(* IEC 61131-3 sources: plc-process-lib/tests/POUs/Suites/FB_Valve_Test (part 2) *)

(* ---- PowerLossStopsWithoutFault.method.impl.st ---- *)
coUnit.TEST('Valve_PowerLoss_StopsWithoutFault');

stCfg.tTravel := T#10S;
fbVlv.xZsc := TRUE;
fbVlv(itfTime := fbTime, stCmd := stCmd, stRetain := stRetain, stCfg := stCfg);
stCmd.xOpen := TRUE;
fbVlv(itfTime := fbTime, stCmd := stCmd, stRetain := stRetain, stCfg := stCfg);
fbVlv.xZsc := FALSE;
FOR iStep := 1 TO 10 DO
    fbTime.Advance(tStep := T#100MS);
    fbVlv(itfTime := fbTime, stCmd := stCmd, stRetain := stRetain, stCfg := stCfg);
END_FOR
fbVlv.xPowerOk := FALSE;
fbTime.Advance(tStep := T#100MS);
fbVlv(itfTime := fbTime, stCmd := stCmd, stRetain := stRetain, stCfg := stCfg);
AssertTrue(Condition := fbVlv.stSts.eState = E_ValveState.Intermediate, Message := 'Intermediate on power loss');
AssertFalse(Condition := fbVlv.xQOpen, Message := 'output off');
AssertEquals_WORD(Expected := GVL_Const.VLV_WRN_POWER_LOST,
                  Actual := fbVlv.stSts.stCommon.wWarning AND GVL_Const.VLV_WRN_POWER_LOST, Message := 'POWER_LOST');
AssertEquals_WORD(Expected := 0, Actual := fbVlv.stSts.stCommon.wFault, Message := 'no fault');
AssertFalse(Condition := fbVlv.Fault, Message := 'not Fault');
stCmd.xOpen := TRUE;
fbTime.Advance(tStep := T#100MS);
fbVlv(itfTime := fbTime, stCmd := stCmd, stRetain := stRetain, stCfg := stCfg);
AssertTrue(Condition := fbVlv.stSts.stCommon.eCmdResult = E_CmdResult.RejectedInhibit,
           Message := 'command without power: RejectedInhibit');
FOR iStep := 1 TO 120 DO                                                // 12 с без напряжения
    fbTime.Advance(tStep := T#100MS);
    fbVlv(itfTime := fbTime, stCmd := stCmd, stRetain := stRetain, stCfg := stCfg);
END_FOR
AssertEquals_WORD(Expected := 0, Actual := fbVlv.stSts.stCommon.wFault, Message := 'travel supervision suspended');
fbVlv.xPowerOk := TRUE;
fbTime.Advance(tStep := T#100MS);
fbVlv(itfTime := fbTime, stCmd := stCmd, stRetain := stRetain, stCfg := stCfg);
AssertTrue(Condition := fbVlv.stSts.eState = E_ValveState.Intermediate, Message := 'Manual stays: target cleared');
AssertFalse(Condition := fbVlv.xQOpen, Message := 'no output in Manual');
stCmd.stCommon.xSetAuto := TRUE;
fbVlv.xAutoOpen := TRUE;
fbTime.Advance(tStep := T#100MS);
fbVlv(itfTime := fbTime, stCmd := stCmd, stRetain := stRetain, stCfg := stCfg);
AssertTrue(Condition := fbVlv.xQOpen, Message := 'Auto drives to target');
AssertTrue(Condition := fbVlv.Available, Message := 'available in Auto with power');
fbVlv.xPowerOk := FALSE;
fbTime.Advance(tStep := T#100MS);
fbVlv(itfTime := fbTime, stCmd := stCmd, stRetain := stRetain, stCfg := stCfg);
AssertFalse(Condition := fbVlv.xQOpen, Message := 'off again without power');
AssertFalse(Condition := fbVlv.Available, Message := 'not available without power');
AssertEquals_WORD(Expected := 0, Actual := fbVlv.stSts.stCommon.wStatus AND GVL_Const.VLV_STS_AVAILABLE,
                  Message := 'AVAILABLE bit off without power');
fbVlv.xPowerOk := TRUE;
fbTime.Advance(tStep := T#100MS);
fbVlv(itfTime := fbTime, stCmd := stCmd, stRetain := stRetain, stCfg := stCfg);
AssertTrue(Condition := fbVlv.xQOpen, Message := 'Auto resumes after power returns');
AssertTrue(Condition := fbVlv.stSts.eState = E_ValveState.Opening, Message := 'Opening');

coUnit.TEST_FINISHED();

(* ---- ResetCauseClearsWithinWindowFaultCleared.method.decl.st ---- *)
// TorqueTrip, Reset при сработавшей муфте: отказ держится; муфта отпустила через 1 с — отказ снят в окне
// tResetWindow без второго результата (и после конца окна RejectedFault нет).
METHOD PRIVATE ResetCauseClearsWithinWindowFaultCleared
VAR
    fbTime   : FB_FakeTime;       // подменное время, старт 1 ч
    fbVlv    : FB_Valve;          // арматура под тестом
    stCmd    : ST_ValveCmd;       // команды HMI
    stRetain : ST_DeviceRetain;   // режим Manual по умолчанию, счётчики
    stCfg    : ST_ValveCfg;       // конфигурация (умолчания: Motorized, ZSO и ZSC)
    iStep    : INT;               // шаг цикла
    uiSeq    : UINT;              // номер команды после Reset
END_VAR

(* ---- ResetCauseClearsWithinWindowFaultCleared.method.impl.st ---- *)
coUnit.TEST('Valve_Reset_CauseClearsWithinWindow_FaultCleared');

stCfg.xTorqueUsed := TRUE;
fbVlv.xZsc := TRUE;
fbVlv(itfTime := fbTime, stCmd := stCmd, stRetain := stRetain, stCfg := stCfg);
stCmd.xOpen := TRUE;
fbVlv(itfTime := fbTime, stCmd := stCmd, stRetain := stRetain, stCfg := stCfg);
fbVlv.xZsc := FALSE;
FOR iStep := 1 TO 10 DO
    fbTime.Advance(tStep := T#100MS);
    fbVlv(itfTime := fbTime, stCmd := stCmd, stRetain := stRetain, stCfg := stCfg);
END_FOR
fbVlv.xTorqueOpen := TRUE;
fbTime.Advance(tStep := T#100MS);
fbVlv(itfTime := fbTime, stCmd := stCmd, stRetain := stRetain, stCfg := stCfg);
AssertEquals_WORD(Expected := GVL_Const.VLV_FLT_TORQUE_TRIP, Actual := fbVlv.stSts.stCommon.wFault,
                  Message := 'TorqueTrip');
stCmd.stCommon.xReset := TRUE;
// t1: Reset, муфта сработана
fbVlv(itfTime := fbTime, stCmd := stCmd, stRetain := stRetain, stCfg := stCfg);
uiSeq := fbVlv.stSts.stCommon.uiCmdSeq;
AssertEquals_WORD(Expected := GVL_Const.VLV_FLT_TORQUE_TRIP, Actual := fbVlv.stSts.stCommon.wFault,
                  Message := 'cause active right after Reset');
FOR iStep := 1 TO 9 DO                                                  // t1 + 0,9 с
    fbTime.Advance(tStep := T#100MS);
    fbVlv(itfTime := fbTime, stCmd := stCmd, stRetain := stRetain, stCfg := stCfg);
END_FOR
AssertEquals_WORD(Expected := GVL_Const.VLV_FLT_TORQUE_TRIP, Actual := fbVlv.stSts.stCommon.wFault,
                  Message := 'still faulted while torque is on');
fbVlv.xTorqueOpen := FALSE;
fbTime.Advance(tStep := T#100MS);
// t1 + 1,0 с: муфта отпустила
fbVlv(itfTime := fbTime, stCmd := stCmd, stRetain := stRetain, stCfg := stCfg);
AssertEquals_WORD(Expected := 0, Actual := fbVlv.stSts.stCommon.wFault, Message := 'cleared within the window');
FOR iStep := 1 TO 30 DO                                                 // дальше конца окна
    fbTime.Advance(tStep := T#100MS);
    fbVlv(itfTime := fbTime, stCmd := stCmd, stRetain := stRetain, stCfg := stCfg);
END_FOR
AssertEquals_UINT(Expected := uiSeq, Actual := fbVlv.stSts.stCommon.uiCmdSeq, Message := 'no second result');
AssertTrue(Condition := fbVlv.stSts.stCommon.eCmdResult = E_CmdResult.Accepted, Message := 'last result Accepted');
AssertFalse(Condition := fbVlv.xQOpen, Message := 'no restart in Manual');

coUnit.TEST_FINISHED();

(* ---- ReverseAfterEndStopWaitsReversePause.method.decl.st ---- *)
// Motorized: ход на открытие дошёл до ZSO на t1 (выход «открывать» снят), сразу команда «закрыть»:
// выход «закрывать» не включается, пока от снятия «открывать» не прошла пауза tReverse = 1 с (на
// t1 + 0,9 с — ещё нет), ровно на t1 + 1,0 с — Closing. То же после стопа в ходе на закрытие (t2) и
// команды «открыть» через 0,2 с: «открывать» включается только на t2 + 1,0 с. Двигатель на выбеге
// встречным включением не реверсируется, даже если ход перед этим остановил концевик или стоп.
METHOD PRIVATE ReverseAfterEndStopWaitsReversePause
VAR
    fbTime   : FB_FakeTime;       // подменное время, старт 1 ч
    fbVlv    : FB_Valve;          // арматура под тестом
    stCmd    : ST_ValveCmd;       // команды HMI
    stRetain : ST_DeviceRetain;   // режим Manual по умолчанию, счётчики
    stCfg    : ST_ValveCfg;       // конфигурация (умолчания: Motorized, ZSO и ZSC, tReverse = 1 с)
    iStep    : INT;               // шаг цикла
    xEverOn  : BOOL;              // выход включался во время паузы
END_VAR

(* ---- ReverseAfterEndStopWaitsReversePause.method.impl.st ---- *)
coUnit.TEST('Valve_ReverseAfterEndStop_WaitsReversePause');

fbVlv.xZsc := TRUE;
// закрыта
fbVlv(itfTime := fbTime, stCmd := stCmd, stRetain := stRetain, stCfg := stCfg);
stCmd.xOpen := TRUE;
fbVlv(itfTime := fbTime, stCmd := stCmd, stRetain := stRetain, stCfg := stCfg);
fbVlv.xZsc := FALSE;
FOR iStep := 1 TO 20 DO                                                 // открывается 2 с
    fbTime.Advance(tStep := T#100MS);
    fbVlv(itfTime := fbTime, stCmd := stCmd, stRetain := stRetain, stCfg := stCfg);
END_FOR
fbVlv.xZso := TRUE;
fbTime.Advance(tStep := T#100MS);
// t1: ZSO, выход «открывать» снят
fbVlv(itfTime := fbTime, stCmd := stCmd, stRetain := stRetain, stCfg := stCfg);
AssertTrue(Condition := fbVlv.stSts.eState = E_ValveState.Open, Message := 'Open on ZSO');
AssertFalse(Condition := fbVlv.xQOpen, Message := 'open contactor off at ZSO');
stCmd.xClose := TRUE;
fbTime.Advance(tStep := T#100MS);
// t1 + 0,1 с: команда «закрыть»
fbVlv(itfTime := fbTime, stCmd := stCmd, stRetain := stRetain, stCfg := stCfg);
AssertTrue(Condition := fbVlv.stSts.stCommon.eCmdResult = E_CmdResult.Accepted, Message := 'close accepted');
xEverOn := fbVlv.xQOpen OR fbVlv.xQClose;
FOR iStep := 1 TO 8 DO                                                  // до t1 + 0,9 с
    fbTime.Advance(tStep := T#100MS);
    fbVlv(itfTime := fbTime, stCmd := stCmd, stRetain := stRetain, stCfg := stCfg);
    xEverOn := xEverOn OR fbVlv.xQOpen OR fbVlv.xQClose;
END_FOR
AssertFalse(Condition := xEverOn, Message := 'no reverse start within tReverse after end stop');
AssertTrue(Condition := fbVlv.stSts.eState = E_ValveState.Open, Message := 'waits at Open');
fbTime.Advance(tStep := T#100MS);
// t1 + 1,0 с
fbVlv(itfTime := fbTime, stCmd := stCmd, stRetain := stRetain, stCfg := stCfg);
AssertTrue(Condition := fbVlv.stSts.eState = E_ValveState.Closing, Message := 'Closing at t1 + tReverse');
AssertTrue(Condition := fbVlv.xQClose, Message := 'close contactor on at t1 + tReverse');
fbVlv.xZso := FALSE;
FOR iStep := 1 TO 20 DO                                                 // закрывается 2 с
    fbTime.Advance(tStep := T#100MS);
    fbVlv(itfTime := fbTime, stCmd := stCmd, stRetain := stRetain, stCfg := stCfg);
END_FOR
stCmd.xStop := TRUE;
// t2: стоп в ходе
fbVlv(itfTime := fbTime, stCmd := stCmd, stRetain := stRetain, stCfg := stCfg);
AssertTrue(Condition := fbVlv.stSts.eState = E_ValveState.Intermediate, Message := 'Intermediate after stop');
stCmd.xOpen := TRUE;
fbTime.Advance(tStep := T#200MS);
// t2 + 0,2 с: команда «открыть»
fbVlv(itfTime := fbTime, stCmd := stCmd, stRetain := stRetain, stCfg := stCfg);
AssertTrue(Condition := fbVlv.stSts.stCommon.eCmdResult = E_CmdResult.Accepted, Message := 'open accepted');
xEverOn := fbVlv.xQOpen OR fbVlv.xQClose;
FOR iStep := 1 TO 7 DO                                                  // до t2 + 0,9 с
    fbTime.Advance(tStep := T#100MS);
    fbVlv(itfTime := fbTime, stCmd := stCmd, stRetain := stRetain, stCfg := stCfg);
    xEverOn := xEverOn OR fbVlv.xQOpen OR fbVlv.xQClose;
END_FOR
AssertFalse(Condition := xEverOn, Message := 'no reverse start within tReverse after stop');
fbTime.Advance(tStep := T#100MS);
// t2 + 1,0 с
fbVlv(itfTime := fbTime, stCmd := stCmd, stRetain := stRetain, stCfg := stCfg);
AssertTrue(Condition := fbVlv.stSts.eState = E_ValveState.Opening, Message := 'Opening at t2 + tReverse');
AssertTrue(Condition := fbVlv.xQOpen, Message := 'open contactor on at t2 + tReverse');

coUnit.TEST_FINISHED();

(* ---- ReversePausesBeforeOppositeDirection.method.decl.st ---- *)
// Motorized открывается; команда «закрыть» в ходе: Reversing, оба выхода сняты на tReverse = 1 с (на
// t1 + 0,9 с ещё сняты), ровно на t1 + 1,0 с включается xQClose.
METHOD PRIVATE ReversePausesBeforeOppositeDirection
VAR
    fbTime   : FB_FakeTime;       // подменное время, старт 1 ч
    fbVlv    : FB_Valve;          // арматура под тестом
    stCmd    : ST_ValveCmd;       // команды HMI
    stRetain : ST_DeviceRetain;   // режим Manual по умолчанию, счётчики
    stCfg    : ST_ValveCfg;       // конфигурация (умолчания: Motorized, ZSO и ZSC)
    iStep    : INT;               // шаг цикла
    xEverOn  : BOOL;              // выход включался во время паузы
END_VAR

(* ---- ReversePausesBeforeOppositeDirection.method.impl.st ---- *)
coUnit.TEST('Valve_Reverse_PausesBeforeOppositeDirection');

fbVlv.xZsc := TRUE;
// закрыта
fbVlv(itfTime := fbTime, stCmd := stCmd, stRetain := stRetain, stCfg := stCfg);
stCmd.xOpen := TRUE;
// Opening
fbVlv(itfTime := fbTime, stCmd := stCmd, stRetain := stRetain, stCfg := stCfg);
fbVlv.xZsc := FALSE;
FOR iStep := 1 TO 20 DO                                                 // открывается 2 с
    fbTime.Advance(tStep := T#100MS);
    fbVlv(itfTime := fbTime, stCmd := stCmd, stRetain := stRetain, stCfg := stCfg);
END_FOR
AssertTrue(Condition := fbVlv.xQOpen, Message := 'opening');
stCmd.xClose := TRUE;
// t1: смена направления
fbVlv(itfTime := fbTime, stCmd := stCmd, stRetain := stRetain, stCfg := stCfg);
AssertTrue(Condition := fbVlv.stSts.eState = E_ValveState.Reversing, Message := 'Reversing on direction change');
AssertFalse(Condition := fbVlv.xQOpen OR fbVlv.xQClose, Message := 'both outputs off during the pause');
AssertTrue(Condition := fbVlv.stSts.stCommon.eCmdResult = E_CmdResult.Accepted, Message := 'close accepted');
FOR iStep := 1 TO 9 DO                                                  // t1 + 0,9 с
    fbTime.Advance(tStep := T#100MS);
    fbVlv(itfTime := fbTime, stCmd := stCmd, stRetain := stRetain, stCfg := stCfg);
    xEverOn := xEverOn OR fbVlv.xQOpen OR fbVlv.xQClose;
END_FOR
AssertFalse(Condition := xEverOn, Message := 'outputs stay off before tReverse');
AssertTrue(Condition := fbVlv.stSts.eState = E_ValveState.Reversing, Message := 'still reversing at t1 + 0.9 s');
fbTime.Advance(tStep := T#100MS);
// t1 + 1,0 с
fbVlv(itfTime := fbTime, stCmd := stCmd, stRetain := stRetain, stCfg := stCfg);
AssertTrue(Condition := fbVlv.stSts.eState = E_ValveState.Closing, Message := 'Closing after tReverse');
AssertTrue(Condition := fbVlv.xQClose, Message := 'close contactor on');
AssertFalse(Condition := fbVlv.xQOpen, Message := 'open contactor off');

coUnit.TEST_FINISHED();

(* ---- SolenoidByTimeCoilOffNotReportedOpen.method.decl.st ---- *)
// Соленоид НЗ (SolenoidEto, без тока закрыт) без концевиков, Manual: открыт по времени хода (tTravel =
// 2 с, катушка под током). Пропало напряжение: катушка без тока, клапан уходит на пружину — «открыто»
// снято (Unknown). Напряжение вернулось: Manual стоит (цель снята), катушка без тока, «открыто» не
// показывается. Снова открыт по времени; Local и возврат в Manual: клапан, закрывшийся на пружине в
// Local, сам не открывается — катушка без команды не включается.
METHOD PRIVATE SolenoidByTimeCoilOffNotReportedOpen
VAR
    fbTime   : FB_FakeTime;       // подменное время, старт 1 ч
    fbVlv    : FB_Valve;          // арматура под тестом
    stCmd    : ST_ValveCmd;       // команды HMI
    stRetain : ST_DeviceRetain;   // режим Manual по умолчанию, счётчики
    stCfg    : ST_ValveCfg;       // конфигурация: SolenoidEto без концевиков
    iStep    : INT;               // шаг цикла
    xEverOn  : BOOL;              // катушка включалась без команды
END_VAR

(* ---- SolenoidByTimeCoilOffNotReportedOpen.method.impl.st ---- *)
coUnit.TEST('Valve_SolenoidByTime_CoilOff_NotReportedOpen');

stCfg.eType := E_ValveType.SolenoidEto;
stCfg.xZsoUsed := FALSE;
stCfg.xZscUsed := FALSE;
stCfg.tTravel := T#2S;
fbVlv(itfTime := fbTime, stCmd := stCmd, stRetain := stRetain, stCfg := stCfg);
stCmd.xOpen := TRUE;
fbVlv(itfTime := fbTime, stCmd := stCmd, stRetain := stRetain, stCfg := stCfg);
FOR iStep := 1 TO 20 DO                                                 // 2 с: открыт по времени
    fbTime.Advance(tStep := T#100MS);
    fbVlv(itfTime := fbTime, stCmd := stCmd, stRetain := stRetain, stCfg := stCfg);
END_FOR
AssertTrue(Condition := fbVlv.stSts.eState = E_ValveState.Open, Message := 'Open by travel time');
AssertTrue(Condition := fbVlv.xQCoil, Message := 'coil holds open');
fbVlv.xPowerOk := FALSE;
fbTime.Advance(tStep := T#100MS);
fbVlv(itfTime := fbTime, stCmd := stCmd, stRetain := stRetain, stCfg := stCfg);
AssertFalse(Condition := fbVlv.xQCoil, Message := 'coil off without power');
AssertFalse(Condition := fbVlv.xOpened, Message := 'spring closes: not reported open');
AssertTrue(Condition := fbVlv.stSts.eState = E_ValveState.Unknown, Message := 'Unknown without coil current');
fbVlv.xPowerOk := TRUE;
fbTime.Advance(tStep := T#100MS);
fbVlv(itfTime := fbTime, stCmd := stCmd, stRetain := stRetain, stCfg := stCfg);
AssertFalse(Condition := fbVlv.xQCoil, Message := 'Manual stays: coil off after power returns');
AssertFalse(Condition := fbVlv.xOpened, Message := 'still not reported open');
stCmd.xOpen := TRUE;
fbVlv(itfTime := fbTime, stCmd := stCmd, stRetain := stRetain, stCfg := stCfg);
FOR iStep := 1 TO 20 DO                                                 // снова открыт по времени
    fbTime.Advance(tStep := T#100MS);
    fbVlv(itfTime := fbTime, stCmd := stCmd, stRetain := stRetain, stCfg := stCfg);
END_FOR
AssertTrue(Condition := fbVlv.stSts.eState = E_ValveState.Open, Message := 'Open by travel time again');
fbVlv.xLocal := TRUE;
fbTime.Advance(tStep := T#100MS);
fbVlv(itfTime := fbTime, stCmd := stCmd, stRetain := stRetain, stCfg := stCfg);
AssertFalse(Condition := fbVlv.xQCoil, Message := 'coil off in Local');
AssertFalse(Condition := fbVlv.xOpened, Message := 'not reported open in Local');
fbVlv.xLocal := FALSE;
FOR iStep := 1 TO 10 DO                                                 // снова Manual, 1 с
    fbTime.Advance(tStep := T#100MS);
    fbVlv(itfTime := fbTime, stCmd := stCmd, stRetain := stRetain, stCfg := stCfg);
    xEverOn := xEverOn OR fbVlv.xQCoil;
END_FOR
AssertTrue(Condition := fbVlv.Mode = E_DeviceMode.Manual, Message := 'back to Manual');
AssertFalse(Condition := xEverOn, Message := 'coil not energized without a command after Local');
AssertFalse(Condition := fbVlv.xOpened, Message := 'not reported open after Local');

coUnit.TEST_FINISHED();

(* ---- SolenoidEtcFaultDeenergizesCoil.method.decl.st ---- *)
// Соленоид НО (SolenoidEtc, без тока открыт): закрытие — катушка под током и держит Closed. Внешняя
// авария — Fault, катушка обесточена (положение пружины, независимо от eSafePos), выходов привода нет;
// причина ушла — катушка без тока до Reset, пружина открыла клапан (xOpened).
METHOD PRIVATE SolenoidEtcFaultDeenergizesCoil
VAR
    fbTime   : FB_FakeTime;       // подменное время, старт 1 ч
    fbVlv    : FB_Valve;          // арматура под тестом
    stCmd    : ST_ValveCmd;       // команды HMI
    stRetain : ST_DeviceRetain;   // режим Manual по умолчанию, счётчики
    stCfg    : ST_ValveCfg;       // конфигурация (умолчания: Motorized, ZSO и ZSC)
    iStep    : INT;               // шаг цикла
END_VAR

(* ---- SolenoidEtcFaultDeenergizesCoil.method.impl.st ---- *)
coUnit.TEST('Valve_SolenoidEtc_FaultDeenergizesCoil');

stCfg.eType := E_ValveType.SolenoidEtc;
fbVlv.xZso := TRUE;
// без тока: открыт
fbVlv(itfTime := fbTime, stCmd := stCmd, stRetain := stRetain, stCfg := stCfg);
AssertTrue(Condition := fbVlv.stSts.eState = E_ValveState.Open, Message := 'normally open valve is Open');
AssertFalse(Condition := fbVlv.xQCoil, Message := 'coil off when open');
stCmd.xClose := TRUE;
fbVlv(itfTime := fbTime, stCmd := stCmd, stRetain := stRetain, stCfg := stCfg);
AssertTrue(Condition := fbVlv.xQCoil, Message := 'coil on to close');
AssertTrue(Condition := fbVlv.stSts.eState = E_ValveState.Closing, Message := 'Closing');
FOR iStep := 1 TO 10 DO
    fbTime.Advance(tStep := T#100MS);
    fbVlv.xZso := FALSE;
    fbVlv.xZsc := iStep >= 10;
    fbVlv(itfTime := fbTime, stCmd := stCmd, stRetain := stRetain, stCfg := stCfg);
END_FOR
AssertTrue(Condition := fbVlv.stSts.eState = E_ValveState.Closed, Message := 'Closed on ZSC');
AssertTrue(Condition := fbVlv.xQCoil, Message := 'coil holds the valve closed');
fbVlv.xExtFault := TRUE;
fbTime.Advance(tStep := T#100MS);
fbVlv(itfTime := fbTime, stCmd := stCmd, stRetain := stRetain, stCfg := stCfg);
AssertFalse(Condition := fbVlv.xQCoil, Message := 'fault: coil de-energized (spring position)');
AssertTrue(Condition := fbVlv.stSts.eState = E_ValveState.Fault, Message := 'Fault');
AssertEquals_WORD(Expected := GVL_Const.VLV_FLT_EXT_FAULT, Actual := fbVlv.stSts.stCommon.wFault,
                  Message := 'wFault ExtFault');
AssertFalse(Condition := fbVlv.xQOpen OR fbVlv.xQClose, Message := 'no motor outputs for a solenoid valve');
fbVlv.xExtFault := FALSE;
fbVlv.xZsc := FALSE;
fbVlv.xZso := TRUE;
fbTime.Advance(tStep := T#100MS);
// пружина открыла клапан
fbVlv(itfTime := fbTime, stCmd := stCmd, stRetain := stRetain, stCfg := stCfg);
AssertFalse(Condition := fbVlv.xQCoil, Message := 'coil stays off until Reset');
AssertTrue(Condition := fbVlv.xOpened, Message := 'spring opened the valve');

coUnit.TEST_FINISHED();

(* ---- SolenoidEtoOpenEnergizesCoil.method.decl.st ---- *)
// Соленоид НЗ (SolenoidEto, без тока закрыт): xOpen — катушка под током, Opening, выходов привода нет;
// ZSO — Open, катушка держит; xClose — катушка обесточена, Closing.
METHOD PRIVATE SolenoidEtoOpenEnergizesCoil
VAR
    fbTime   : FB_FakeTime;       // подменное время, старт 1 ч
    fbVlv    : FB_Valve;          // арматура под тестом
    stCmd    : ST_ValveCmd;       // команды HMI
    stRetain : ST_DeviceRetain;   // режим Manual по умолчанию, счётчики
    stCfg    : ST_ValveCfg;       // конфигурация (умолчания: Motorized, ZSO и ZSC)
    iStep    : INT;               // шаг цикла
END_VAR

(* ---- SolenoidEtoOpenEnergizesCoil.method.impl.st ---- *)
coUnit.TEST('Valve_SolenoidEto_OpenEnergizesCoil');

stCfg.eType := E_ValveType.SolenoidEto;
fbVlv.xZsc := TRUE;
fbVlv(itfTime := fbTime, stCmd := stCmd, stRetain := stRetain, stCfg := stCfg);
AssertFalse(Condition := fbVlv.xQCoil, Message := 'coil off when closed');
stCmd.xOpen := TRUE;
fbVlv(itfTime := fbTime, stCmd := stCmd, stRetain := stRetain, stCfg := stCfg);
AssertTrue(Condition := fbVlv.xQCoil, Message := 'coil energized to open');
AssertTrue(Condition := fbVlv.stSts.eState = E_ValveState.Opening, Message := 'Opening');
AssertFalse(Condition := fbVlv.xQOpen OR fbVlv.xQClose, Message := 'no motor outputs');
FOR iStep := 1 TO 10 DO
    fbTime.Advance(tStep := T#100MS);
    fbVlv.xZsc := FALSE;
    fbVlv.xZso := iStep >= 10;
    fbVlv(itfTime := fbTime, stCmd := stCmd, stRetain := stRetain, stCfg := stCfg);
END_FOR
AssertTrue(Condition := fbVlv.stSts.eState = E_ValveState.Open, Message := 'Open on ZSO');
AssertTrue(Condition := fbVlv.xQCoil, Message := 'coil holds the valve open');
stCmd.xClose := TRUE;
fbTime.Advance(tStep := T#100MS);
fbVlv(itfTime := fbTime, stCmd := stCmd, stRetain := stRetain, stCfg := stCfg);
AssertFalse(Condition := fbVlv.xQCoil, Message := 'coil off to close');
AssertTrue(Condition := fbVlv.stSts.eState = E_ValveState.Closing, Message := 'Closing');

coUnit.TEST_FINISHED();

(* ---- SolenoidWithZsoPowerLossNoPositionLostFault.method.decl.st ---- *)
// Соленоидный клапан НЗ (SolenoidEto) с ZSO и ZSC, открыт командой до ZSO. Пропало питание привода: катушка
// обесточена, клапан уходит на пружину — ZSO пропал, через 1 с ZSC. Отказа PositionLost нет: без напряжения уход
// с концевика не контролируется (VLV-08), состояние Closed. Питание вернулось — отказа нет, в Manual катушка не
// включается.
METHOD PRIVATE SolenoidWithZsoPowerLossNoPositionLostFault
VAR
    fbTime   : FB_FakeTime;       // подменное время, старт 1 ч
    fbVlv    : FB_Valve;          // арматура под тестом
    stCmd    : ST_ValveCmd;       // команды HMI
    stRetain : ST_DeviceRetain;   // режим, счётчики
    stCfg    : ST_ValveCfg;       // конфигурация (умолчания: Motorized, ZSO и ZSC)
    iStep    : INT;               // шаг цикла

    wFltSeen : WORD;              // отказы, которые хоть раз появлялись
END_VAR

(* ---- SolenoidWithZsoPowerLossNoPositionLostFault.method.impl.st ---- *)
coUnit.TEST('Valve_SolenoidWithZso_PowerLoss_NoPositionLostFault');

stCfg.eType := E_ValveType.SolenoidEto;
fbVlv.xZsc := TRUE;
fbVlv(itfTime := fbTime, stCmd := stCmd, stRetain := stRetain, stCfg := stCfg);   // t0: Closed по ZSC
stCmd.xOpen := TRUE;
fbTime.Advance(tStep := T#100MS);
fbVlv(itfTime := fbTime, stCmd := stCmd, stRetain := stRetain, stCfg := stCfg);   // Opening, катушка
fbVlv.xZsc := FALSE;
fbVlv.xZso := TRUE;
fbTime.Advance(tStep := T#100MS);
fbVlv(itfTime := fbTime, stCmd := stCmd, stRetain := stRetain, stCfg := stCfg);   // Open по ZSO
AssertTrue(Condition := fbVlv.xQCoil AND fbVlv.stSts.eState = E_ValveState.Open,
           Message := 'precondition: open on ZSO, coil holds');
fbVlv.xPowerOk := FALSE;
fbTime.Advance(tStep := T#100MS);
fbVlv(itfTime := fbTime, stCmd := stCmd, stRetain := stRetain, stCfg := stCfg);       // нет напряжения
fbVlv.xZso := FALSE;                                                                   // пружина
FOR iStep := 1 TO 10 DO
    fbTime.Advance(tStep := T#100MS);
    fbVlv(itfTime := fbTime, stCmd := stCmd, stRetain := stRetain, stCfg := stCfg);
    wFltSeen := wFltSeen OR fbVlv.stSts.stCommon.wFault;
END_FOR
fbVlv.xZsc := TRUE;
fbTime.Advance(tStep := T#100MS);
fbVlv(itfTime := fbTime, stCmd := stCmd, stRetain := stRetain, stCfg := stCfg);       // ZSC
AssertEquals_WORD(Expected := 0, Actual := wFltSeen OR fbVlv.stSts.stCommon.wFault,
                  Message := 'no PositionLost without power');
AssertTrue(Condition := fbVlv.stSts.eState = E_ValveState.Closed, Message := 'Closed by ZSC');
AssertFalse(Condition := fbVlv.xQCoil, Message := 'coil off');
fbVlv.xPowerOk := TRUE;
FOR iStep := 1 TO 10 DO
    fbTime.Advance(tStep := T#100MS);
    fbVlv(itfTime := fbTime, stCmd := stCmd, stRetain := stRetain, stCfg := stCfg);
END_FOR
AssertEquals_WORD(Expected := 0, Actual := fbVlv.stSts.stCommon.wFault, Message := 'no fault after power returns');
AssertFalse(Condition := fbVlv.xQCoil, Message := 'Manual: no output after power returns');

coUnit.TEST_FINISHED();

(* ---- StopMotorizedGoesIntermediate.method.decl.st ---- *)
// Motorized открывается; xStop в ходе — Intermediate, выходы сняты, Accepted, бит сброшен. Цель Manual
// «никуда»: арматура стоит и дальше.
METHOD PRIVATE StopMotorizedGoesIntermediate
VAR
    fbTime   : FB_FakeTime;       // подменное время, старт 1 ч
    fbVlv    : FB_Valve;          // арматура под тестом
    stCmd    : ST_ValveCmd;       // команды HMI
    stRetain : ST_DeviceRetain;   // режим Manual по умолчанию, счётчики
    stCfg    : ST_ValveCfg;       // конфигурация (умолчания: Motorized, ZSO и ZSC)
    iStep    : INT;               // шаг цикла
    xEverOn  : BOOL;              // выход включался после стопа
END_VAR

(* ---- StopMotorizedGoesIntermediate.method.impl.st ---- *)
coUnit.TEST('Valve_StopMotorized_GoesIntermediate');

fbVlv.xZsc := TRUE;
fbVlv(itfTime := fbTime, stCmd := stCmd, stRetain := stRetain, stCfg := stCfg);
stCmd.xOpen := TRUE;
fbVlv(itfTime := fbTime, stCmd := stCmd, stRetain := stRetain, stCfg := stCfg);
fbVlv.xZsc := FALSE;
FOR iStep := 1 TO 20 DO                                                 // открывается 2 с
    fbTime.Advance(tStep := T#100MS);
    fbVlv(itfTime := fbTime, stCmd := stCmd, stRetain := stRetain, stCfg := stCfg);
END_FOR
stCmd.xStop := TRUE;
fbVlv(itfTime := fbTime, stCmd := stCmd, stRetain := stRetain, stCfg := stCfg);
AssertTrue(Condition := fbVlv.stSts.eState = E_ValveState.Intermediate, Message := 'Intermediate after stop');
AssertFalse(Condition := fbVlv.xQOpen OR fbVlv.xQClose, Message := 'outputs off');
AssertTrue(Condition := fbVlv.stSts.stCommon.eCmdResult = E_CmdResult.Accepted, Message := 'stop accepted');
AssertFalse(Condition := stCmd.xStop, Message := 'xStop cleared');
FOR iStep := 1 TO 20 DO
    fbTime.Advance(tStep := T#100MS);
    fbVlv(itfTime := fbTime, stCmd := stCmd, stRetain := stRetain, stCfg := stCfg);
    xEverOn := xEverOn OR fbVlv.xQOpen OR fbVlv.xQClose;
END_FOR
AssertFalse(Condition := xEverOn, Message := 'stays stopped');
AssertFalse(Condition := fbVlv.xOpened OR fbVlv.xClosed, Message := 'neither open nor closed');

coUnit.TEST_FINISHED();

(* ---- StopSolenoidRejected.method.decl.st ---- *)
// Соленоид НЗ (SolenoidEto) открывается; xStop — RejectedNotSupported: катушка и движение не меняются,
// бит сброшен.
METHOD PRIVATE StopSolenoidRejected
VAR
    fbTime   : FB_FakeTime;       // подменное время, старт 1 ч
    fbVlv    : FB_Valve;          // арматура под тестом
    stCmd    : ST_ValveCmd;       // команды HMI
    stRetain : ST_DeviceRetain;   // режим Manual по умолчанию, счётчики
    stCfg    : ST_ValveCfg;       // конфигурация (умолчания: Motorized, ZSO и ZSC)
END_VAR

(* ---- TorqueMidTravelLatchesTorqueTrip.method.decl.st ---- *)
// Муфта подключена. Через 3 с хода, до концевика, сработала муфта открытия — TorqueTrip (wFault бит 4),
// выход снят, бит TORQUE. Муфта отпустила — отказ держится (бит TORQUE снят); Reset снимает отказ,
// арматура в промежутке стоит (Manual).
METHOD PRIVATE TorqueMidTravelLatchesTorqueTrip
VAR
    fbTime   : FB_FakeTime;       // подменное время, старт 1 ч
    fbVlv    : FB_Valve;          // арматура под тестом
    stCmd    : ST_ValveCmd;       // команды HMI
    stRetain : ST_DeviceRetain;   // режим Manual по умолчанию, счётчики
    stCfg    : ST_ValveCfg;       // конфигурация (умолчания: Motorized, ZSO и ZSC)
    iStep    : INT;               // шаг цикла
END_VAR

(* ---- TorqueMidTravelLatchesTorqueTrip.method.impl.st ---- *)
coUnit.TEST('Valve_TorqueMidTravel_LatchesTorqueTrip');

stCfg.xTorqueUsed := TRUE;
fbVlv.xZsc := TRUE;
fbVlv(itfTime := fbTime, stCmd := stCmd, stRetain := stRetain, stCfg := stCfg);
stCmd.xOpen := TRUE;
fbVlv(itfTime := fbTime, stCmd := stCmd, stRetain := stRetain, stCfg := stCfg);
fbVlv.xZsc := FALSE;
FOR iStep := 1 TO 30 DO                                                 // открывается 3 с
    fbTime.Advance(tStep := T#100MS);
    fbVlv(itfTime := fbTime, stCmd := stCmd, stRetain := stRetain, stCfg := stCfg);
END_FOR
fbVlv.xTorqueOpen := TRUE;
fbTime.Advance(tStep := T#100MS);
// муфта раньше концевика
fbVlv(itfTime := fbTime, stCmd := stCmd, stRetain := stRetain, stCfg := stCfg);
AssertTrue(Condition := fbVlv.stSts.eState = E_ValveState.Fault, Message := 'Fault on torque mid travel');
AssertEquals_WORD(Expected := GVL_Const.VLV_FLT_TORQUE_TRIP, Actual := fbVlv.stSts.stCommon.wFault,
                  Message := 'wFault TorqueTrip');
AssertFalse(Condition := fbVlv.xQOpen, Message := 'output off');
AssertEquals_WORD(Expected := GVL_Const.VLV_STS_TORQUE,
                  Actual := fbVlv.stSts.stCommon.wStatus AND GVL_Const.VLV_STS_TORQUE, Message := 'TORQUE bit');
fbVlv.xTorqueOpen := FALSE;
fbTime.Advance(tStep := T#100MS);
fbVlv(itfTime := fbTime, stCmd := stCmd, stRetain := stRetain, stCfg := stCfg);
AssertEquals_WORD(Expected := GVL_Const.VLV_FLT_TORQUE_TRIP, Actual := fbVlv.stSts.stCommon.wFault,
                  Message := 'latched after the switch released');
AssertEquals_WORD(Expected := 0, Actual := fbVlv.stSts.stCommon.wStatus AND GVL_Const.VLV_STS_TORQUE,
                  Message := 'TORQUE bit follows the switch');
stCmd.stCommon.xReset := TRUE;
fbVlv(itfTime := fbTime, stCmd := stCmd, stRetain := stRetain, stCfg := stCfg);
AssertEquals_WORD(Expected := 0, Actual := fbVlv.stSts.stCommon.wFault, Message := 'cleared by Reset');
AssertTrue(Condition := fbVlv.stSts.eState = E_ValveState.Intermediate, Message := 'Intermediate after Reset');
AssertFalse(Condition := fbVlv.xQOpen, Message := 'no restart in Manual');

coUnit.TEST_FINISHED();
